// TIA Portal V19 export
// export: ExportSetting WithDefaults
Screen "CO_0000_100_Traceability_01"  1920x966, Number=100, Template=CC_0000_ScreenTemplate
  on ClearScreen: SetTag(Tag := Menu_BrowserScreenNo, Value := 0)
  on GenerateScreen: MenuManagement_VB(BrowserScreenNo := Menu_BrowserScreenNoGroup02_Subgroup06)
  ScreenLayer 
    Button "btnLegend" at 1784,3 size 135x81  Mode=Text, TextOff="Leyenda / Legend / Legende", TextOn="Leyenda / Legend / Legende"
      on Release: ShowPopupScreen(Name of the screen := Legend_1201_Traceability_Popup, X coordinate := 760, Y coordinate := 162, Display mode := -1, Animation := 2, Animation speed := 0)
    Button "btnInterlock" at 1647,3 size 135x81  Mode=Text, TextOff="Enclavamiento / Interlock / Verriegelung", TextOn="Enclavamiento / Interlock / Verriegelung"
      on Release: ShowPopupScreen(Name of the screen := Traceability_1203_Interlock_Popup, X coordinate := 860, Y coordinate := 162, Display mode := -1, Animation := 2, Animation speed := 0)
    Button "btnI4.0" at 1510,3 size 135x81  Mode=Text, TextOff="I4.0", TextOn="I4.0"
      RangeAppearanceAnimation "RangeAppearanceAnimation"
        tag I40_Systems_Status
        0..0: back #636571, fore #000000
        1..1: back #00ff00, fore #000000
      on Press: SetBit(Tag := I40_Systems_Reset)
      on Release: ResetBit(Tag := I40_Systems_Reset)
  ScreenLayer 
    FaceplateInstance "fpScreenLocking" at 0,0 size 1920x964  FaceplateTypeName=#SICAR@GST_Types_HMI@$@00_General@$@ScreenLocking V 4.0.0
      on Release_LockedScreen: ShowPopupScreen(Name of the screen := Dialog_BlockedScreen_Popup, X coordinate := 1020, Y coordinate := 162, Display mode := -1, Animation := 2, Animation speed := 1)
      on Release_StopRTPLCConnection: ShowPopupScreen(Name of the screen := Dialog_0801_Settings_StopRuntime_Popup, X coordinate := 1058, Y coordinate := 88, Display mode := 1, Animation := 2, Animation speed := 0); SetTag(Tag := WinccRT_Stop_Selected, Value := 0)
      on Release_StopRTPLCStop: ShowPopupScreen(Name of the screen := Dialog_0801_Settings_StopRuntime_Popup, X coordinate := 1058, Y coordinate := 88, Display mode := 1, Animation := 2, Animation speed := 0); SetTag(Tag := WinccRT_Stop_Selected, Value := 0)
      Connection_State := Connection_state
      PLC_Mode := PlcMode
      Locked_Screen := Menu_ActiveScreenLocked
  ScreenLayer 
    Line "linLineHeader" at 0,86 size 1920x0
    TextField "txtTitleScreen" at 585,3 size 750x40  Text="Trazabilidad / Traceability / Nachvollziehbarkeit"
    SymbolicIOField "outSubtitleScreen" at 686,45 size 549x40  CountVisibleItems=8, Mode=Output, OnValue=1, TextList=CO_Traceability_ID, TextOff="0", TextOn="1"
      ProcessValue := Int_Value_001
